(* IEC 61131-3 sources: model-first-plc-agent-ai/results/T4-W-21, 2 files *)

(* ---- a1_code.st ---- *)
FUNCTION_BLOCK LevelControlRuntime
VAR_INPUT
    StartCommand : BOOL;
    StopCommand : BOOL;
    LevelMeter : INT;
    FULL_SCALE : INT;
    h_sp : REAL;
    h_max : REAL;
    eps : REAL;
    t_h : TIME;
    Kp : REAL;
    Ti : REAL;
    Td : REAL;
    CycleTime : TIME;
END_VAR
VAR_OUTPUT
    FillValve : INT := 0;
    DischargeValve : INT := 0;
    fill_valve : BOOL := FALSE;
    discharge_valve : BOOL := FALSE;
END_VAR
VAR
    StartEdge : R_TRIG;
    HoldTimer : TON;
    start : BOOL;
    stop : BOOL;
    settled : BOOL := FALSE;

    (* Region encoding: 0 = LOW, 1 = MID, 2 = HIGH. *)
    r : INT := 0;

    (* Initial GRAFCET situation: {x0}. *)
    x0 : BOOL := TRUE;
    x1 : BOOL := FALSE;

    h : REAL;
    e : REAL;
    SampleSeconds : REAL;
    IntegralValue : REAL := 0.0;
    IntegralCandidate : REAL;
    PreviousError : REAL := 0.0;
    DerivativeValue : REAL;
    ProportionalValue : REAL;
    RawDemand : REAL;
    BoundedDemand : REAL;
    PidWasActive : BOOL := FALSE;
END_VAR

StartEdge(CLK := StartCommand);
start := StartEdge.Q;
stop := StopCommand;

h := INT_TO_REAL(LevelMeter) / INT_TO_REAL(FULL_SCALE);
e := h_sp - h;

IF h < h_sp THEN
    r := 0;
ELSIF h < h_max THEN
    r := 1;
ELSE
    r := 2;
END_IF;

(* Qualify continuous residence in the tolerance band during x1. *)
HoldTimer(
    IN := x1 AND (ABS(e) <= eps) AND NOT stop,
    PT := t_h
);
settled := HoldTimer.Q;

(* Evaluate only transitions enabled by the preceding situation. *)
IF x0 THEN
    IF start AND NOT stop AND NOT (r = 2) THEN
        x0 := FALSE;
        x1 := TRUE;
    END_IF;
ELSIF x1 THEN
    IF stop OR settled OR (r = 2) THEN
        x1 := FALSE;
        x0 := TRUE;
    END_IF;
END_IF;

(* Non-stored GRAFCET actions. *)
fill_valve := x1;
discharge_valve := x1;

IF NOT x1 THEN
    HoldTimer(IN := FALSE, PT := t_h);
    settled := FALSE;
END_IF;

FillValve := 0;
DischargeValve := 0;

IF fill_valve THEN
    SampleSeconds := TIME_TO_REAL(CycleTime) / 1000.0;

    (* Reset PID state at each new regulation interval. *)
    IF NOT PidWasActive THEN
        IntegralValue := 0.0;
        PreviousError := e;
    END_IF;

    ProportionalValue := Kp * e;
    DerivativeValue := 0.0;

    IF (SampleSeconds > 0.0) AND (Td > 0.0) THEN
        DerivativeValue :=
            Kp * Td * (e - PreviousError) / SampleSeconds;
    END_IF;

    IntegralCandidate := IntegralValue;
    IF (SampleSeconds > 0.0) AND (Ti > 0.0) THEN
        IntegralCandidate :=
            IntegralValue + Kp * e * SampleSeconds / Ti;
    END_IF;

    RawDemand :=
        ProportionalValue + IntegralCandidate + DerivativeValue;

    (* Reject this scan's integral update if it causes saturation. *)
    IF (RawDemand >= 0.0) AND (RawDemand <= 1.0) THEN
        IntegralValue := IntegralCandidate;
    END_IF;

    RawDemand :=
        ProportionalValue + IntegralValue + DerivativeValue;

    IF RawDemand < 0.0 THEN
        BoundedDemand := 0.0;
    ELSIF RawDemand > 1.0 THEN
        BoundedDemand := 1.0;
    ELSE
        BoundedDemand := RawDemand;
    END_IF;

    FillValve :=
        REAL_TO_INT(BoundedDemand * INT_TO_REAL(FULL_SCALE));
    PreviousError := e;
ELSE
    IntegralValue := 0.0;
    PreviousError := e;
END_IF;

IF discharge_valve THEN
    DischargeValve := REAL_TO_INT(0.4 * INT_TO_REAL(FULL_SCALE));
END_IF;

PidWasActive := fill_valve;

END_FUNCTION_BLOCK

PROGRAM Main
VAR
    StartCommand AT %IX100.0 : BOOL;
    StopCommand AT %IX100.1 : BOOL;
    LevelMeter AT %IW100 : INT;
    FillValve AT %QW100 : INT;
    DischargeValve AT %QW101 : INT;
END_VAR
VAR CONSTANT
    FULL_SCALE : INT := 1000;
END_VAR
VAR
    Controller : LevelControlRuntime;

    (* Normalized measuring span: 1.0 corresponds to 10 V. *)
    h_sp : REAL := 0.8;
    h_max : REAL := 0.9;
    eps : REAL := 0.02;
    t_h : TIME := T#10s;

    (* Commissioning parameters; Ti and Td are expressed in seconds. *)
    Kp : REAL := 1.0;
    Ti : REAL := 10.0;
    Td : REAL := 0.0;

    (* Configure the OpenPLC cyclic task to match this period. *)
    CycleTime : TIME := T#20ms;
END_VAR

Controller(
    StartCommand := StartCommand,
    StopCommand := StopCommand,
    LevelMeter := LevelMeter,
    FULL_SCALE := FULL_SCALE,
    h_sp := h_sp,
    h_max := h_max,
    eps := eps,
    t_h := t_h,
    Kp := Kp,
    Ti := Ti,
    Td := Td,
    CycleTime := CycleTime
);

FillValve := Controller.FillValve;
DischargeValve := Controller.DischargeValve;

END_PROGRAM

(* ---- a2_code.st ---- *)
FUNCTION_BLOCK LevelControl
VAR_INPUT
    StartCommand : BOOL;
    StopCommand : BOOL;
    LevelMeter : INT;
    Kp : REAL := 20.0;
    Ti : REAL := 5.0;
    Td : REAL := 0.0;
END_VAR
VAR_OUTPUT
    FillValve : INT;
    DischargeValve : INT;
    fill_valve : BOOL;
    discharge_valve : BOOL;
END_VAR
VAR CONSTANT
    FULL_SCALE : INT := 1000;
    h_span : REAL := 10.0;
    h_sp : REAL := 8.0;
    h_target : REAL := 8.0;
    h_max : REAL := 9.0;
    eps : REAL := 0.2;
    t_h : TIME := T#10s;
    scan_seconds : REAL := 0.02;
    region_low : INT := 0;
    region_middle : INT := 1;
    region_high : INT := 2;
END_VAR
VAR
    start_edge : R_TRIG;
    hold_timer : TON;
    start : BOOL;
    stop : BOOL;
    settled : BOOL;
    r : INT;
    sequence_state : INT := 0;
    x0 : BOOL;
    x1 : BOOL;
    h : REAL;
    e : REAL;
    previous_error : REAL := 0.0;
    integral_term : REAL := 0.0;
    proposed_integral : REAL;
    proportional_term : REAL;
    derivative_term : REAL;
    raw_demand : REAL;
    bounded_demand : REAL;
    pid_initialized : BOOL := FALSE;
END_VAR

(* This block must execute once every 20 ms. Ti and Td are in seconds;
   Kp is in percent valve opening per volt of level error. *)
start_edge(CLK := StartCommand);
start := start_edge.Q;
stop := StopCommand;

h := INT_TO_REAL(LevelMeter) * h_span / INT_TO_REAL(FULL_SCALE);
e := h_sp - h;

IF h < h_target THEN
    r := region_low;
ELSIF h < h_max THEN
    r := region_middle;
ELSE
    r := region_high;
END_IF;

(* The hold condition measures uninterrupted time in the tolerance band,
   and is reset outside regulation or whenever the band is left. *)
hold_timer(
    IN := (sequence_state = 1) AND
          NOT stop AND
          (r <> region_high) AND
          (ABS(e) <= eps),
    PT := t_h
);
settled := hold_timer.Q;

IF stop THEN
    sequence_state := 0;
ELSE
    CASE sequence_state OF
        0:
            IF start AND (r <> region_high) THEN
                sequence_state := 1;
            END_IF;
        1:
            IF settled OR (r = region_high) THEN
                sequence_state := 0;
            END_IF;
    ELSE
        sequence_state := 0;
    END_CASE;
END_IF;

x0 := sequence_state = 0;
x1 := sequence_state = 1;

fill_valve := x1;
discharge_valve := x1;

FillValve := 0;
DischargeValve := 0;

IF fill_valve THEN
    IF NOT pid_initialized THEN
        integral_term := 0.0;
        previous_error := e;
        pid_initialized := TRUE;
    END_IF;

    proportional_term := Kp * e;
    derivative_term := Kp * Td * (e - previous_error) / scan_seconds;

    proposed_integral := integral_term;
    IF Ti > 0.0 THEN
        proposed_integral :=
            integral_term + Kp * e * scan_seconds / Ti;
    ELSE
        (* A nonpositive Ti disables the integral component. *)
        integral_term := 0.0;
        proposed_integral := 0.0;
    END_IF;

    raw_demand :=
        proportional_term + proposed_integral + derivative_term;

    (* Suspend integration whenever the proposed output is clamped. *)
    IF raw_demand > 100.0 THEN
        bounded_demand := 100.0;
    ELSIF raw_demand < 0.0 THEN
        bounded_demand := 0.0;
    ELSE
        bounded_demand := raw_demand;
        integral_term := proposed_integral;
    END_IF;

    previous_error := e;
    FillValve := REAL_TO_INT(
        bounded_demand * INT_TO_REAL(FULL_SCALE) / 100.0
    );
ELSE
    pid_initialized := FALSE;
    integral_term := 0.0;
    previous_error := e;
    bounded_demand := 0.0;
END_IF;

IF discharge_valve THEN
    DischargeValve := REAL_TO_INT(0.4 * INT_TO_REAL(FULL_SCALE));
END_IF;

END_FUNCTION_BLOCK

PROGRAM Main
VAR
    StartCommand AT %IX100.0 : BOOL;
    StopCommand AT %IX100.1 : BOOL;
    LevelMeter AT %IW100 : INT;
    FillValve AT %QW100 : INT;
    DischargeValve AT %QW101 : INT;
END_VAR
VAR
    controller : LevelControl;
    Kp : REAL := 20.0;
    Ti : REAL := 5.0;
    Td : REAL := 0.0;
END_VAR

controller(
    StartCommand := StartCommand,
    StopCommand := StopCommand,
    LevelMeter := LevelMeter,
    Kp := Kp,
    Ti := Ti,
    Td := Td
);

FillValve := controller.FillValve;
DischargeValve := controller.DischargeValve;

END_PROGRAM

CONFIGURATION Config0
    RESOURCE Res0 ON PLC
        TASK ControlTask(INTERVAL := T#20ms, PRIORITY := 0);
        PROGRAM MainInstance WITH ControlTask : Main;
    END_RESOURCE
END_CONFIGURATION
